(* IEC 61131-3 sources: plc-iiot-stack/tests/POUs/FB_JsonBuilder_Test, 11 files *)

(* ---- BufferHoldsExactlyItsSize.method.decl.st ---- *)
// Объект ровно на размер буфера — полный, на байт больше — переполнение.
METHOD PRIVATE BufferHoldsExactlyItsSize
VAR_INST
    fbJson : FB_JsonBuilder;
END_VAR
VAR
    iField : INT;
END_VAR

(* ---- BufferHoldsExactlyItsSize.method.impl.st ---- *)
coUnit.TEST('BufferHoldsExactlyItsSize');

// поле "kkk":"<63 символа>" — 71 байт; «{» и 14 полей с запятыми — 1 + 14 * 71 + 13 = 1008 байт
fbJson.Begin();
FOR iField := 1 TO 14 DO
    fbJson.AddString(sKey := 'kkk', sValue := '123456789012345678901234567890123456789012345678901234567890123');
END_FOR
fbJson.AddString(sKey := 'q', sValue := '1234567');   // ,"q":"1234567" — 14 байт: 1022, «}» — 1023
AssertTrue(Condition := fbJson.Finish(), Message := 'object of exactly the buffer size must fit');
AssertEquals_UINT(Expected := 1023, Actual := fbJson.uiLen, Message := 'length equals buffer size');
fbJson.Begin();
FOR iField := 1 TO 14 DO
    fbJson.AddString(sKey := 'kkk', sValue := '123456789012345678901234567890123456789012345678901234567890123');
END_FOR
fbJson.AddString(sKey := 'q', sValue := '12345678');
AssertFalse(Condition := fbJson.Finish(), Message := 'one byte more must overflow');

coUnit.TEST_FINISHED();

(* ---- BuildsFlatObjectWithAllTypes.method.decl.st ---- *)
// Объект со строкой, целым, логическим, null и числом — точный текст.
METHOD PRIVATE BuildsFlatObjectWithAllTypes
VAR_INST
    fbJson : FB_JsonBuilder;
END_VAR

(* ---- EmptyObjectAndRestart.method.decl.st ---- *)
// Пустой объект; Begin очищает предыдущий текст.
METHOD PRIVATE EmptyObjectAndRestart
VAR_INST
    fbJson : FB_JsonBuilder;
END_VAR

(* ---- EscapesSpecialCharacters.method.decl.st ---- *)
// Экранирование кавычки, обратной косой черты и управляющих символов.
METHOD PRIVATE EscapesSpecialCharacters
VAR_INST
    fbJson : FB_JsonBuilder;
END_VAR

(* ---- IntExtremes.method.decl.st ---- *)
// Целые: 0, максимум и минимум LINT, отметка времени в мс.
METHOD PRIVATE IntExtremes
VAR_INST
    fbJson : FB_JsonBuilder;
END_VAR

(* ---- NotFiniteBecomesNull.method.decl.st ---- *)
// NaN, бесконечность и слишком большие числа пишутся как null.
METHOD PRIVATE NotFiniteBecomesNull
VAR_INST
    fbJson : FB_JsonBuilder;
END_VAR
VAR
    lwNan : LWORD := 16#7FF8000000000000;
    lwInf : LWORD := 16#7FF0000000000000;
    pBits : POINTER TO LREAL;
    lrNan : LREAL;
    lrInf : LREAL;
END_VAR

(* ---- OverflowIsReportedNotTruncatedSilently.method.decl.st ---- *)
// Переполнение буфера: xOverflow, Finish = FALSE, длина не больше буфера.
METHOD PRIVATE OverflowIsReportedNotTruncatedSilently
VAR_INST
    fbJson : FB_JsonBuilder;
END_VAR
VAR
    iField : INT;
END_VAR

(* ---- OverflowIsReportedNotTruncatedSilently.method.impl.st ---- *)
coUnit.TEST('OverflowIsReportedNotTruncatedSilently');

fbJson.Begin();
FOR iField := 1 TO 40 DO
    fbJson.AddString(sKey := 'key_with_some_length', sValue := 'value with some length to fill the buffer');
END_FOR
AssertFalse(Condition := fbJson.Finish(), Message := 'Finish must fail after overflow');
AssertTrue(Condition := fbJson.xOverflow, Message := 'overflow flag must be set');
AssertEquals_UINT(Expected := GVL_Const.MQTT_PAYLOAD_LEN, Actual := fbJson.uiLen,
                  Message := 'buffer is filled up to its size and not beyond');

coUnit.TEST_FINISHED();

(* ---- RealFormattingRoundsAndTrimsZeros.method.decl.st ---- *)
// Числа: округление до знаков, без хвостовых нулей, -0 как 0, предел знаков.
METHOD PRIVATE RealFormattingRoundsAndTrimsZeros
VAR_INST
    fbJson : FB_JsonBuilder;
END_VAR

(* ---- RealFromRealIsRoundedLikeTheValueShown.method.decl.st ---- *)
// REAL 2.35 (в двоичном виде 2.3499999) с тремя знаками — 2.35.
METHOD PRIVATE RealFromRealIsRoundedLikeTheValueShown
VAR_INST
    fbJson : FB_JsonBuilder;
END_VAR
VAR
    rValue : REAL := 2.35;
END_VAR
